// High-rate recording chunk — struct-of-arrays (SoA) so the app can bulk-read
// each channel as a flat typed array over ADS (no struct packing/alignment).
//
// One CHUNK = REC_CHUNK EtherCAT frames. The recorder FB fills the active chunk
// one frame per cycle; when full it advances to the next chunk in the ring and
// bumps GVL_Recording.nChunkSeq. The app reads each completed chunk's arrays in
// one bulk ADS read per channel, then writes them to the recording file.
//
// Two rates share one DC timebase:
//   * bus-rate  (one value per frame): aDcTs + load motors / Futek / Mentee status
//   * Mentee    (REC_OVERSAMPLE per frame): aMn* arrays, length REC_CHUNK*REC_OVERSAMPLE
//
// Sizes are compile-time constants in GVL_Recording — keep them in lock-step
// with the FB and the backend reader (chunk length + oversample count).
TYPE ST_RecChunk :
STRUCT
    nCount   : UDINT;   // frames actually filled in this chunk (= REC_CHUNK when complete)

    // ── bus-rate channels (one element per frame) ──────────────────────
    // Types match the source snapshot fields exactly (no implicit conversion):
    // load motors / analog are LREAL; encoder counters are DWORD.
    aDcTs    : ARRAY[0..GVL_Recording.REC_CHUNK - 1] OF ULINT;   // DC time, 100 ns ticks
    aM1Pos   : ARRAY[0..GVL_Recording.REC_CHUNK - 1] OF LREAL;   // load motor 1
    aM1Vel   : ARRAY[0..GVL_Recording.REC_CHUNK - 1] OF LREAL;
    aM1Trq   : ARRAY[0..GVL_Recording.REC_CHUNK - 1] OF LREAL;
    aM2Pos   : ARRAY[0..GVL_Recording.REC_CHUNK - 1] OF LREAL;   // load motor 2
    aM2Vel   : ARRAY[0..GVL_Recording.REC_CHUNK - 1] OF LREAL;
    aM2Trq   : ARRAY[0..GVL_Recording.REC_CHUNK - 1] OF LREAL;
    aEnc1Cnt : ARRAY[0..GVL_Recording.REC_CHUNK - 1] OF DWORD;   // Futek 1 encoder
    aEnc1Frq : ARRAY[0..GVL_Recording.REC_CHUNK - 1] OF DWORD;
    aEnc2Cnt : ARRAY[0..GVL_Recording.REC_CHUNK - 1] OF DWORD;   // Futek 2 encoder
    aEnc2Frq : ARRAY[0..GVL_Recording.REC_CHUNK - 1] OF DWORD;
    aAin1V   : ARRAY[0..GVL_Recording.REC_CHUNK - 1] OF LREAL;   // Futek 1 analog (V)
    aAin2V   : ARRAY[0..GVL_Recording.REC_CHUNK - 1] OF LREAL;   // Futek 2 analog (V)
    aMnSW    : ARRAY[0..GVL_Recording.REC_CHUNK - 1] OF UDINT;   // Mentee status word (bus-rate)
    aMnCnt   : ARRAY[0..GVL_Recording.REC_CHUNK - 1] OF UDINT;   // fresh oversamples this frame (0..REC_OVERSAMPLE)

    // ── Mentee oversamples (REC_OVERSAMPLE per frame) — raw slot words ──
    // w0/w1/w2 are raw 32-bit words for the fixed lanes (theta / d_theta / iq).
    // Storing them raw keeps the recorder decode-agnostic — the app reinterprets
    // the bits per lane.
    aMnIdx   : ARRAY[0..GVL_Recording.REC_CHUNK * GVL_Recording.REC_OVERSAMPLE - 1] OF UDINT; // sample_idx
    aMnW0    : ARRAY[0..GVL_Recording.REC_CHUNK * GVL_Recording.REC_OVERSAMPLE - 1] OF UDINT;
    aMnW1    : ARRAY[0..GVL_Recording.REC_CHUNK * GVL_Recording.REC_OVERSAMPLE - 1] OF UDINT;
    aMnW2    : ARRAY[0..GVL_Recording.REC_CHUNK * GVL_Recording.REC_OVERSAMPLE - 1] OF UDINT;
    // ── extended lanes 3..9 — ELF-picked debug variables (slot-2 pipe) ──
    // Same flat index as aMnIdx/aMnW0..2 (frame*REC_OVERSAMPLE + slot), so
    // element i of EVERY aMn* array is the same synchronized capture instant.
    // Kept LAST so the app can skip reading them when nothing is selected.
    aMnW3    : ARRAY[0..GVL_Recording.REC_CHUNK * GVL_Recording.REC_OVERSAMPLE - 1] OF UDINT;
    aMnW4    : ARRAY[0..GVL_Recording.REC_CHUNK * GVL_Recording.REC_OVERSAMPLE - 1] OF UDINT;
    aMnW5    : ARRAY[0..GVL_Recording.REC_CHUNK * GVL_Recording.REC_OVERSAMPLE - 1] OF UDINT;
    aMnW6    : ARRAY[0..GVL_Recording.REC_CHUNK * GVL_Recording.REC_OVERSAMPLE - 1] OF UDINT;
    aMnW7    : ARRAY[0..GVL_Recording.REC_CHUNK * GVL_Recording.REC_OVERSAMPLE - 1] OF UDINT;
    aMnW8    : ARRAY[0..GVL_Recording.REC_CHUNK * GVL_Recording.REC_OVERSAMPLE - 1] OF UDINT;
    aMnW9    : ARRAY[0..GVL_Recording.REC_CHUNK * GVL_Recording.REC_OVERSAMPLE - 1] OF UDINT;

    // ── Futek analog oversamples (REC_FUTEK_OS per frame) — EL3702 x5, in Volts ──
    // Flat index frame*REC_FUTEK_OS + slot. Stored as V (same scale as aAin1V) so
    // the backend's volts->Nm calibration path handles them identically, at 5x rate.
    aFut1V   : ARRAY[0..GVL_Recording.REC_CHUNK * GVL_Recording.REC_FUTEK_OS - 1] OF LREAL;   // Futek 1 (stAnalogIn1 ch1)
    aFut2V   : ARRAY[0..GVL_Recording.REC_CHUNK * GVL_Recording.REC_FUTEK_OS - 1] OF LREAL;   // Futek 2 (stAnalogIn2 ch1)
END_STRUCT
END_TYPE

(* stored: Version 1.1.0.1, ProductVersion 3.1.4026.18
   DUT ST_RecChunk: Id {a1f4c7e2-1d33-4b8a-9c64-7e2a5f1b9d40} *)
